(* IEC 61131-3 sources: llm-plc-st-eval/data/processed_v2_primera/gpt-4o/B2/few_shot, 3 files *)

(* ---- ejec_1.st ---- *)
FUNCTION_BLOCK FB_Valvula
VAR_INPUT
    nivelAlto : BOOL; (* Sensor de nivel alto *)
END_VAR
VAR_OUTPUT
    valvula : BOOL; (* Válvula de drenaje *)
END_VAR
VAR
    tRetardo : TON; (* Temporizador de retardo *)
END_VAR

(* La válvula se abre si el nivel alto se mantiene durante 5 segundos *)
tRetardo(IN := nivelAlto, PT := T#5S);
valvula := tRetardo.Q;
END_FUNCTION_BLOCK

(* ---- ejec_2.st ---- *)
FUNCTION_BLOCK FB_Valvula
VAR_INPUT
    nivelAlto : BOOL; (* Sensor de nivel alto *)
END_VAR
VAR_OUTPUT
    valvula : BOOL; (* Válvula de drenaje *)
END_VAR
VAR
    tRetardo : TON; (* Temporizador de retardo *)
END_VAR

(* La válvula se abre si el nivel alto se mantiene durante 5 segundos *)
tRetardo(IN := nivelAlto, PT := T#5S);
valvula := tRetardo.Q;
END_FUNCTION_BLOCK

(* ---- ejec_3.st ---- *)
FUNCTION_BLOCK FB_Valvula
VAR_INPUT
    nivelAlto : BOOL; (* Sensor de nivel alto *)
END_VAR
VAR_OUTPUT
    valvula : BOOL; (* Válvula de drenaje *)
END_VAR
VAR
    tRetardo : TON; (* Temporizador de retardo *)
END_VAR

(* La válvula se abre si el nivel alto se mantiene durante 5 segundos *)
tRetardo(IN := nivelAlto, PT := T#5S);
valvula := tRetardo.Q;
END_FUNCTION_BLOCK
